(* PLC project c.project, CODESYS CODESYS V3.5 SP17 Patch 3 *)
(* stored: creationDateTime 2026-10-19T00:00:00, modificationDateTime 2026-10-19T00:00:00 *)

PROGRAM PRG_S
VAR_INPUT
    go : BOOL;
END_VAR
VAR_OUTPUT
    n : INT;
END_VAR

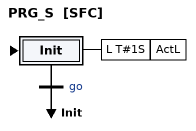
INITIAL_STEP Init:
  ActL(L, T#1S);
END_STEP
TRANSITION FROM Init TO Init
  := go;
END_TRANSITION

ACTION ActL:
                n := n + 1;

              
END_ACTION
END_PROGRAM
